(*
SPDX-FileCopyrightText: © 2026 Oleksandr Tiutyk <trofimich@gmail.com>
SPDX-License-Identifier: MIT
License: https://opensource.org/license/mit
*)

(*!
<summary>
Beckhoff PWM output channel process image.
</summary>
<description>
Represents the duty-only EL2502 standard PWM PDO with signed presentation selected through CoE.
DutyCycle 0..32767 represents 0..100 percent before user scaling; frequency is configured acyclically.
Cyclic-period and unsigned-presentation variants are outside this channel. No clamping or CoE configuration occurs.
When used for I/O, link located fields or their containing buffers to the matching selected PDOs.
The record is not a packed wire buffer; compiler padding is not part of the device specification.
Unlinked/default values do not prove valid I/O. The caller evaluates bus/channel validity before use.
Use one owner task per instance and externally synchronize other access; multi-field snapshots are not atomic.
Copies store data without creating hardware links. Keep borrowed field references valid while consumers are bound.
This passive record performs no validation, synchronization, configuration or protocol advancement.
</description>
*)
TYPE PWM_OUTPUT_CHANNEL :
STRUCT
	DutyCycle AT %Q* : INT;
END_STRUCT
END_TYPE

(* stored: Version 1.1.0.1, ProductVersion 3.1.4026.20
   DUT PWM_OUTPUT_CHANNEL: Id {d2e58131-b13f-4bf4-82f1-5275b3d92441} *)
